
// ===== library: MasterCopy "FB_FIR_LowPass" =====

// folder: UUT/FIR

FUNCTION_BLOCK "FB_FIR_LowPass"   // FB23, SCL
{ S7_Optimized_Access := 'TRUE' }
VERSION : 0.1
   VAR_INPUT
      Enable : Bool;   // filter active
      Reset : Bool;   // restart: the filter is filled with the current X (no start-up ramp)
      X : LReal;   // input sample
      Fc_Set : LReal := 1.0;   // [Hz] requested -3 dB cutoff, about 0.23 Hz ... 20 Hz; a change restarts the filter
      Ts_Limit : LReal := 0.01;   // [s] longer intervals (e.g. a communication peak) are ignored
      Ts_Tol : LReal := 0.05;   // allowed deviation of the average cycle from TS_DESIGN (0.05 = 5 %)
   END_VAR
   VAR_OUTPUT
      Y : LReal;   // filtered output
      M_Act : Int;   // window length of each stage in samples
      Fc_Eff : LReal;   // effective -3 dB cutoff for M_Act and Ts_Meas [Hz]
      Delay : LReal;   // delay of the output (group delay) [s]
      Ts_Meas : LReal;   // average sample period = average OB1 cycle, over about 1 s [s]
      Ts_Valid : Bool;   // TRUE = RUNTIME gave a plausible interval in this call
      Ts_Drift : Bool;   // TRUE = the average cycle differs from TS_DESIGN by more than Ts_Tol: the cutoff is off
   END_VAR
   VAR
      RtMem : LReal;   // memory of RUNTIME
      First : Bool := TRUE;   // first call: no interval yet
      HaveTs : Bool;   // TRUE after the first valid interval
      TsAvg : LReal;   // average of the valid intervals [s]
      Filled : Bool;   // TRUE after the buffers were filled
      "M" : Int;   // window length in use
      Pos : Int;   // ring buffer index: oldest sample of every stage, overwritten in this call
      Sum : Array[0..3] of LReal;   // running sum of every stage
      Buf : Array[0..3, 0..999] of LReal;   // last M inputs of every stage; second bound = M_MAX - 1
   END_VAR
   VAR_TEMP
      tsRaw : LReal;
      mReq : DInt;
      v : LReal;
      s : Int;
      i : Int;
   END_VAR
   VAR CONSTANT
      STAGE_LAST : Int := 3;   // 4 stages
      M_MAX : Int := 1000;   // bound of #Buf: lowest cutoff about 0.23 Hz at 1 ms
      TS_DESIGN : LReal := 0.001;   // design sample period = OB1 cycle [s]
      FC_FACTOR : LReal := 0.2276;   // 4 stages: -3 dB cutoff = FC_FACTOR / (M * Ts)
      TS_SMOOTH : LReal := 0.001;   // weight of a new interval in #TsAvg (about 1000 cycles = 1 s)
   END_VAR
BEGIN

    REGION Description
        // FIR low-pass made of 4 cascaded moving averages of M samples each (4 * (M - 1) + 1 taps, all positive):
        // linear phase, DC gain 1, no overshoot on a step. Every stage keeps a running sum, so one call costs the
        // same for any M: the cutoff can go low without more computing time, only more memory (#Buf).
        //   -3 dB at Fc = 0.2276 / (M * Ts); zeros at multiples of 1 / (M * Ts); everything above the first zero
        //   is damped by at least 53 dB. Delay = 2 * (M - 1) * Ts, about 0.45 / Fc.
        // M follows from Fc_Set and TS_DESIGN (rounded, 1 ... M_MAX), so Fc_Eff differs slightly from Fc_Set.
        // Call in every OB1 cycle and unconditionally: RUNTIME measures the time between two calls.
    END_REGION

    REGION Sample period (RUNTIME: time since the previous call, in seconds)
        #tsRaw := RUNTIME(#RtMem);
        #Ts_Valid := NOT #First AND #tsRaw > 0.0 AND #tsRaw <= #Ts_Limit;
        #First := FALSE;
        IF #Ts_Valid THEN
            IF #HaveTs THEN
                #TsAvg := #TsAvg + (#tsRaw - #TsAvg) * #TS_SMOOTH;
            ELSE
                #TsAvg := #tsRaw;
                #HaveTs := TRUE;
            END_IF;
        END_IF;
        // an invalid interval keeps the last average; before the first valid one: design period
        IF #HaveTs THEN
            #Ts_Meas := #TsAvg;
        ELSE
            #Ts_Meas := #TS_DESIGN;
        END_IF;
        #Ts_Drift := #HaveTs AND ABS(#Ts_Meas - #TS_DESIGN) > #Ts_Tol * #TS_DESIGN;
    END_REGION

    REGION Window length from the requested cutoff
        // LREAL_TO_DINT rounds to the nearest value; below the lowest cutoff: M_MAX (also for Fc_Set <= 0)
        IF #Fc_Set > #FC_FACTOR / (INT_TO_LREAL(#M_MAX) * #TS_DESIGN) THEN
            #mReq := LREAL_TO_DINT(#FC_FACTOR / (#Fc_Set * #TS_DESIGN));
        ELSE
            #mReq := INT_TO_DINT(#M_MAX);
        END_IF;
        IF #mReq < 1 THEN
            #mReq := 1;
        END_IF;
    END_REGION

    REGION Filter
        IF #Reset OR NOT #Filled OR #mReq <> INT_TO_DINT(#M) THEN
            // (re)start: fill every stage with the current input, so the output starts at X
            #M := DINT_TO_INT(#mReq);
            FOR #s := 0 TO #STAGE_LAST DO
                FOR #i := 0 TO #M - 1 DO
                    #Buf[#s, #i] := #X;
                END_FOR;
                #Sum[#s] := #X * INT_TO_LREAL(#M);
            END_FOR;
            #Pos := 0;
            #Filled := TRUE;
            #Y := #X;
        ELSIF #Enable THEN
            #v := #X;
            FOR #s := 0 TO #STAGE_LAST DO
                #Sum[#s] := #Sum[#s] + #v - #Buf[#s, #Pos];   // add the newest, drop the oldest
                #Buf[#s, #Pos] := #v;
                #v := #Sum[#s] / INT_TO_LREAL(#M);   // average of this stage = input of the next one
            END_FOR;
            #Pos := #Pos + 1;
            IF #Pos >= #M THEN
                #Pos := 0;
            END_IF;
            #Y := #v;
        END_IF;

        #M_Act := #M;
        #Fc_Eff := #FC_FACTOR / (INT_TO_LREAL(#M) * #Ts_Meas);
        #Delay := 2.0 * INT_TO_LREAL(#M - 1) * #Ts_Meas;
    END_REGION
END_FUNCTION_BLOCK

// ===== library: MasterCopy "FB_FIR_LP100" =====

// folder: UUT/FIR

FUNCTION_BLOCK "FB_FIR_LP100"   // FB21, SCL
{ S7_Optimized_Access := 'TRUE' }
VERSION : 0.4
   VAR_INPUT
      Enable : Bool;   // filter active
      Reset : Bool;   // clear the delay line
      X : LReal;   // input sample
      Ts_Limit : LReal := 0.01;   // [s] longer intervals (e.g. a communication peak) are ignored
      Ts_Tol : LReal := 0.05;   // allowed deviation of the average cycle from TS_DESIGN (0.05 = 5 %)
   END_VAR
   VAR_OUTPUT
      Y : LReal;   // filtered output
      Ts_Meas : LReal;   // average sample period = average OB1 cycle, over about 1 s [s]
      Ts_Valid : Bool;   // TRUE = RUNTIME gave a plausible interval in this call
      Ts_Drift : Bool;   // TRUE = the average cycle differs from TS_DESIGN by more than Ts_Tol: the cutoff is off
      Fc_Eff : LReal;   // effective -3 dB cutoff for Ts_Meas [Hz]
   END_VAR
   VAR
      RtMem : LReal;   // memory of RUNTIME
      First : Bool := TRUE;   // first call: no interval yet
      HaveTs : Bool;   // TRUE after the first valid interval
      TsAvg : LReal;   // average of the valid intervals [s]
      Pos : Int;   // index of the newest sample in #Line (ring buffer)
      Line : Array[0..16] of LReal;   // delay line (ring buffer)
      Coef : Array[0..16] of LReal;   // [0] [1] [2] [3] [4] [5] [6] [7] [8] [9] [10] [11] [12] [13] [14] [15] [16] filter taps, do not change online
   END_VAR
   VAR_TEMP
      tsRaw : LReal;
      acc : LReal;
      i : Int;
      j : Int;
   END_VAR
   VAR CONSTANT
      LAST_TAP : Int := 16;   // number of taps - 1 = upper bound of #Line and #Coef
      TS_DESIGN : LReal := 0.001;   // design sample period = OB1 cycle [s], fs = 1000 Hz
      FC_DESIGN : LReal := 100.0;   // design -3 dB cutoff [Hz]
      TS_SMOOTH : LReal := 0.001;   // weight of a new interval in #TsAvg (about 1000 cycles = 1 s)
   END_VAR
   // Coef[0] := -1.48651536431772E-19;
   // Coef[1] := -0.000353560113498742;
   // Coef[2] := -0.00350832878720326;
   // Coef[3] := -0.00907130526178393;
   // Coef[4] := -0.00367490473275513;
   // Coef[5] := 0.037817961535658;
   // Coef[6] := 0.124770149738866;
   // Coef[7] := 0.221633438427618;
   // Coef[8] := 0.264773098386197;
   // Coef[9] := 0.221633438427618;
   // Coef[10] := 0.124770149738866;
   // Coef[11] := 0.037817961535658;
   // Coef[12] := -0.00367490473275513;
   // Coef[13] := -0.00907130526178392;
   // Coef[14] := -0.00350832878720326;
   // Coef[15] := -0.000353560113498744;
   // Coef[16] := -1.48651536431772E-19;
BEGIN

    REGION Description
        // FIR low-pass, 17 taps (Blackman-windowed sinc), linear phase, group delay 8 samples = 8 ms, DC gain 1.
        // Designed for an OB1 cycle of 1 ms: -3 dB at 100 Hz, -60 dB from 287 Hz, below -72 dB from 300 Hz to 500 Hz.
        // The taps are fixed, so the cutoff scales with the average cycle: Fc_Eff = 100 Hz * TS_DESIGN / Ts_Meas.
        // Ts_Drift reports a lasting deviation; short peaks of the cycle are averaged out.
        // Call in every OB1 cycle and unconditionally: RUNTIME measures the time between two calls.
    END_REGION

    REGION Sample period (RUNTIME: time since the previous call, in seconds)
        #tsRaw := RUNTIME(#RtMem);
        #Ts_Valid := NOT #First AND #tsRaw > 0.0 AND #tsRaw <= #Ts_Limit;
        #First := FALSE;
        IF #Ts_Valid THEN
            IF #HaveTs THEN
                #TsAvg := #TsAvg + (#tsRaw - #TsAvg) * #TS_SMOOTH;
            ELSE
                #TsAvg := #tsRaw;
                #HaveTs := TRUE;
            END_IF;
        END_IF;
        // an invalid interval keeps the last average; before the first valid one: design period
        IF #HaveTs THEN
            #Ts_Meas := #TsAvg;
        ELSE
            #Ts_Meas := #TS_DESIGN;
        END_IF;
        #Fc_Eff := #FC_DESIGN * #TS_DESIGN / #Ts_Meas;
        #Ts_Drift := #HaveTs AND ABS(#Ts_Meas - #TS_DESIGN) > #Ts_Tol * #TS_DESIGN;
    END_REGION

    REGION Convolution (ring buffer: one write per cycle instead of shifting all samples)
        IF #Reset THEN
            FOR #i := 0 TO #LAST_TAP DO
                #Line[#i] := 0.0;
            END_FOR;
            #Pos := 0;
            #Y := 0.0;
        ELSIF #Enable THEN
            #Pos := #Pos + 1;
            IF #Pos > #LAST_TAP THEN
                #Pos := 0;
            END_IF;
            #Line[#Pos] := #X;
            #acc := 0.0;
            #j := #Pos;   // Coef[i] * sample of i cycles ago
            FOR #i := 0 TO #LAST_TAP DO
                #acc := #acc + #Coef[#i] * #Line[#j];
                #j := #j - 1;
                IF #j < 0 THEN
                    #j := #LAST_TAP;
                END_IF;
            END_FOR;
            #Y := #acc;
        END_IF;
    END_REGION
END_FUNCTION_BLOCK

// ===== library: MasterCopy "UnitTest_FIR_LowPass" =====

// folder: UUT/FIR

FUNCTION_BLOCK "UnitTest_FIR_LowPass"   // FB22, SCL
{ S7_Optimized_Access := 'TRUE' }
VERSION : 0.1
   VAR_INPUT
      reset : Bool;   // TRUE = start the test again (as "DB_UnitTestControl".reset)
   END_VAR
   VAR_OUTPUT
      Done : Bool;   // TRUE when all test steps are finished
   END_VAR
   VAR_IN_OUT
      "Step" : UDInt;   // current step; only increases: 0, 10, 20, 30, 40, 9900
   END_VAR
   VAR
      TestCase : String[24];   // signal of the current step (online monitoring)
      Fir : "FB_FIR_LowPass";   // device under test
      StepTimer : TON_TIME;   // 5 s per signal
      StepRun : Bool;   // FALSE for one cycle after a step change: restarts #StepTimer
      StepSamples : DInt;   // filter calls since the start of the step
      Counting : Bool;   // TRUE = the filter has settled and, for a sine, a signal period has started
      Seed : DWord := 16#2545_F491;   // state of the noise generator (xorshift32), never 0; restarted in step 0
      Sig : Struct   // signal of the current step: X = Offset + Amp * sin(Phase) + noise
         Offset : LReal;
         Amp : LReal;
         K : LReal;   // frequency as a multiple of the effective cutoff: f = K * Fc_Eff
         NoiseAmp : LReal;   // uniform noise in -NoiseAmp ... +NoiseAmp
         FreqHz : LReal;   // resulting frequency (online monitoring)
         Phase : LReal;
         Noise : LReal;
         X : LReal;   // filter input
      END_STRUCT;
      Acc : Struct   // running sums while #Counting
         N : DInt;
         SumY : LReal;
         SumY2 : LReal;
         SumI : LReal;   // Y * sin(Phase)
         SumQ : LReal;   // Y * cos(Phase)
      END_STRUCT;
      Full : Struct   // sums of #Acc at the end of the last whole signal period (sine steps)
         N : DInt;
         SumI : LReal;
         SumQ : LReal;
      END_STRUCT;
      Result : Array[1..4] of Struct   // one entry per signal step: measured value and limits
         Value : LReal;   // step 10: mean of Y; steps 20 ... 40: amplitude of Y at the signal frequency
         Lo : LReal;
         Hi : LReal;
         N : DInt;   // evaluated samples; 0 = the step was too short for an evaluation
         Pass : Bool;
      END_STRUCT;
      NoiseRatio : LReal;   // step 10: standard deviation of Y / standard deviation of the input noise
   END_VAR
   VAR_TEMP
      _ret : Bool;
      res : Int;   // index into #Result
      mean : LReal;
   END_VAR
   VAR CONSTANT
      LAST_STEP : UDInt := 16#FFFF_FFFF;
      STEP_FINISH : UDInt := 9900;
      STEP_TIME : Time := T#5S;   // duration of every signal
      TEST_FC : LReal := 10.0;   // [Hz] cutoff under test: M = 11, so the slow sine of step 20 fits into 5 s
      TWO_PI : LReal := 6.28318530717959;
      NOISE_RATIO_MAX : LReal := 0.3;   // white noise gain of the taps for M = 11 is 0.209
   END_VAR
BEGIN

    REGION BLOCK INFO HEADER
        //===============================================================================
        // Title:            Unit test for FB_FIR_LowPass
        // Comment/Function: Four signals with uniform noise, 5 s each; checks DC gain, noise reduction,
        //                   passband, -3 dB point and stopband at Fc_Set = TEST_FC
        // Requirements:     "FB_FIR_LowPass", unit test framework ("BeforeEach", "AfterEach", "assertTrue",
        //                   "DB_UnitTestControl")
        // Restrictions:     call in every OB1 cycle, unconditionally. The OB1 cycle must be below about 4 ms,
        //                   otherwise 5 s give too few samples (step 10 and step 20 become unreliable)
        //-------------------------------------------------------------------------------
        // Change log table:
        // Version  | Date       | Expert in charge       | Changes applied
        //----------|------------|------------------------|------------------------------
        // 00.00.01 | 21.11.2026 | Roman Butsenko
        //                         First released version, from UnitTest_FIR_LP100 V0.0.3
        //===============================================================================
    END_REGION
    REGION Description
        // Steps (each signal runs STEP_TIME; the evaluation starts after the filter length, 4 * M_Act calls):
        //   10  DC 1.0 + noise 0.5     -> mean of Y 0.98 ... 1.02, noise std reduced below NOISE_RATIO_MAX
        //   20  sine 0.1 * Fc + noise  -> amplitude 0.95 ... 1.05 (passband, theory 0.997)
        //   30  sine 1.0 * Fc + noise  -> amplitude 0.65 ... 0.76 (-3 dB point, theory 0.707)
        //   40  sine 6.6 * Fc + noise  -> amplitude <= 0.004 (stopband, 1.5 x first zero, theory 0.0023 = -53 dB)
        // The filter runs with Fc_Set = TEST_FC; M only scales the filter, so other cutoffs behave the same.
        // Fc is "Fir".Fc_Eff, so the signal has the same frequency per filter call for any OB1 cycle. The amplitude
        // is measured by correlation with sin and cos of the signal phase over whole signal periods, which ignores
        // the noise and the filter delay. Results: #Result[1..4], #NoiseRatio.
    END_REGION

    REGION Reset
        IF "DB_UnitTestControl".reset = 1 OR #reset THEN
            #Done := FALSE;
            #Step := 0;
            #StepRun := FALSE;
            #TestCase := '';
            RETURN;
        END_IF;
    END_REGION

    REGION Signal of this step
        CASE #Step OF
            10:
                #TestCase := 'DC + noise';
                #Sig.Offset := 1.0; #Sig.Amp := 0.0; #Sig.K := 0.0; #Sig.NoiseAmp := 0.5;
            20:
                #TestCase := 'Sine 0.1 Fc + noise';
                #Sig.Offset := 0.0; #Sig.Amp := 1.0; #Sig.K := 0.1; #Sig.NoiseAmp := 0.2;
            30:
                #TestCase := 'Sine 1.0 Fc + noise';
                #Sig.Offset := 0.0; #Sig.Amp := 1.0; #Sig.K := 1.0; #Sig.NoiseAmp := 0.2;
            40:
                #TestCase := 'Sine 6.6 Fc + noise';
                #Sig.Offset := 0.0; #Sig.Amp := 1.0; #Sig.K := 6.6; #Sig.NoiseAmp := 0.2;
            ELSE
                #Sig.Offset := 0.0; #Sig.Amp := 0.0; #Sig.K := 0.0; #Sig.NoiseAmp := 0.0;
        END_CASE;

        // noise: xorshift32, scaled to -NoiseAmp ... +NoiseAmp
        #Seed := #Seed XOR SHL(IN := #Seed, N := 13);
        #Seed := #Seed XOR SHR(IN := #Seed, N := 17);
        #Seed := #Seed XOR SHL(IN := #Seed, N := 5);
        #Sig.Noise := (UDINT_TO_LREAL(DWORD_TO_UDINT(#Seed)) / 4294967296.0 * 2.0 - 1.0) * #Sig.NoiseAmp;
        #Sig.X := #Sig.Offset + #Sig.Amp * SIN(#Sig.Phase) + #Sig.Noise;

        #Fir(Enable := TRUE,
             Reset := #Step = 0,
             X := #Sig.X,
             Fc_Set := #TEST_FC);
        #StepSamples := #StepSamples + 1;

        // step timer: restarts one cycle after every step change
        #StepTimer(IN := #StepRun, PT := #STEP_TIME);
        #StepRun := TRUE;

        // running sums
        IF #Counting THEN
            #Acc.N := #Acc.N + 1;
            #Acc.SumY := #Acc.SumY + #Fir.Y;
            #Acc.SumY2 := #Acc.SumY2 + #Fir.Y * #Fir.Y;
            #Acc.SumI := #Acc.SumI + #Fir.Y * SIN(#Sig.Phase);
            #Acc.SumQ := #Acc.SumQ + #Fir.Y * COS(#Sig.Phase);
        END_IF;

        // next phase: f = K * Fc_Eff; Fc_Eff * Ts_Meas is constant, so the phase step per call is constant
        #Sig.FreqHz := #Sig.K * #Fir.Fc_Eff;
        #Sig.Phase := #Sig.Phase + #TWO_PI * #Sig.FreqHz * #Fir.Ts_Meas;
        IF #Sig.Phase >= #TWO_PI THEN   // a signal period is complete
            #Sig.Phase := #Sig.Phase - #TWO_PI;
            IF #Counting THEN   // keep the sums over whole periods
                #Full.N := #Acc.N;
                #Full.SumI := #Acc.SumI;
                #Full.SumQ := #Acc.SumQ;
            ELSIF #StepSamples >= 4 * INT_TO_DINT(#Fir.M_Act) THEN   // settled: start counting with a new period
                #Counting := TRUE;
            END_IF;
        END_IF;
        IF #Sig.K = 0.0 AND #StepSamples >= 4 * INT_TO_DINT(#Fir.M_Act) THEN   // DC: no periods, count once settled
            #Counting := TRUE;
        END_IF;
    END_REGION

    REGION Test steps
        CASE #Step OF
            0:
                "BeforeEach"(iName := GetBlockName(DINT#16));
                #Result[1].Lo := 0.98;  #Result[1].Hi := 1.02;
                #Result[2].Lo := 0.95;  #Result[2].Hi := 1.05;
                #Result[3].Lo := 0.65;  #Result[3].Hi := 0.76;
                #Result[4].Lo := 0.0;   #Result[4].Hi := 0.004;
                #NoiseRatio := 0.0;
                #Seed := 16#2545_F491;   // same noise in every run, so a failure can be repeated
                #Step := 10;
                #StepRun := FALSE;
                #StepSamples := 0;
                #Counting := FALSE;
                #Sig.Phase := 0.0;
                #Acc.N := 0; #Acc.SumY := 0.0; #Acc.SumY2 := 0.0; #Acc.SumI := 0.0; #Acc.SumQ := 0.0;
                #Full.N := 0; #Full.SumI := 0.0; #Full.SumQ := 0.0;

            10, 20, 30, 40:
                IF #StepTimer.Q THEN
                    #res := UDINT_TO_INT(#Step / 10);
                    #Result[#res].Value := 0.0;
                    IF #Step = 10 THEN
                        #Result[#res].N := #Acc.N;
                        IF #Acc.N > 0 THEN
                            #mean := #Acc.SumY / DINT_TO_LREAL(#Acc.N);
                            #Result[#res].Value := #mean;
                            // std of Y / std of the input noise (uniform: NoiseAmp / sqrt(3))
                            #NoiseRatio := SQRT(MAX(IN1 := #Acc.SumY2 / DINT_TO_LREAL(#Acc.N) - #mean * #mean, IN2 := 0.0))
                                           / (#Sig.NoiseAmp / SQRT(3.0));
                            #_ret := "assertTrue"(#NoiseRatio <= #NOISE_RATIO_MAX);   // noise is reduced
                        END_IF;
                    ELSE
                        #Result[#res].N := #Full.N;
                        IF #Full.N > 0 THEN
                            #Result[#res].Value := 2.0 / DINT_TO_LREAL(#Full.N) * SQRT(#Full.SumI * #Full.SumI + #Full.SumQ * #Full.SumQ);
                        END_IF;
                    END_IF;
                    #Result[#res].Pass := #Result[#res].N > 0 AND #Result[#res].Value >= #Result[#res].Lo AND #Result[#res].Value <= #Result[#res].Hi;
                    #_ret := "assertTrue"(#Result[#res].Pass);

                    // next signal
                    IF #Step < 40 THEN
                        #Step := #Step + 10;
                    ELSE
                        #Step := #STEP_FINISH;
                    END_IF;
                    #StepRun := FALSE;
                    #StepSamples := 0;
                    #Counting := FALSE;
                    #Sig.Phase := 0.0;
                    #Acc.N := 0; #Acc.SumY := 0.0; #Acc.SumY2 := 0.0; #Acc.SumI := 0.0; #Acc.SumQ := 0.0;
                    #Full.N := 0; #Full.SumI := 0.0; #Full.SumQ := 0.0;
                END_IF;

            #STEP_FINISH: // all test steps are done
                #Done := TRUE;
                "AfterEach"();
                #Step := #LAST_STEP;

            #LAST_STEP:
                // just idle
                ;

            ELSE // step number without a label: report it and finish the test
                #_ret := "assertTrue"(FALSE);
                #Step := #STEP_FINISH;
        END_CASE;
    END_REGION
END_FUNCTION_BLOCK

// ===== library: MasterCopy "UnitTest_FIR_LP100" =====

// folder: UUT/FIR

FUNCTION_BLOCK "UnitTest_FIR_LP100"   // FB20, SCL
{ S7_Optimized_Access := 'TRUE' }
VERSION : 0.3
   VAR_INPUT
      reset : Bool;   // TRUE = start the test again (as "DB_UnitTestControl".reset)
   END_VAR
   VAR_OUTPUT
      Done : Bool;   // TRUE when all test steps are finished
   END_VAR
   VAR_IN_OUT
      "Step" : UDInt;   // current step; only increases: 0, 10, 20, 30, 40, 9900
   END_VAR
   VAR
      TestCase : String[24];   // signal of the current step (online monitoring)
      Fir : "FB_FIR_LP100";   // device under test
      StepTimer : TON_TIME;   // 5 s per signal
      StepRun : Bool;   // FALSE for one cycle after a step change: restarts #StepTimer
      StepSamples : DInt;   // filter calls since the start of the step
      Counting : Bool;   // TRUE = the filter has settled and, for a sine, a signal period has started
      Seed : DWord := 16#2545_F491;   // state of the noise generator (xorshift32), never 0; restarted in step 0
      Sig : Struct   // signal of the current step: X = Offset + Amp * sin(Phase) + noise
         Offset : LReal;
         Amp : LReal;
         K : LReal;   // frequency as a multiple of the effective cutoff: f = K * Fc_Eff
         NoiseAmp : LReal;   // uniform noise in -NoiseAmp ... +NoiseAmp
         FreqHz : LReal;   // resulting frequency (online monitoring)
         Phase : LReal;
         Noise : LReal;
         X : LReal;   // filter input
      END_STRUCT;
      Acc : Struct   // running sums while #Counting
         N : DInt;
         SumY : LReal;
         SumY2 : LReal;
         SumI : LReal;   // Y * sin(Phase)
         SumQ : LReal;   // Y * cos(Phase)
      END_STRUCT;
      Full : Struct   // sums of #Acc at the end of the last whole signal period (sine steps)
         N : DInt;
         SumI : LReal;
         SumQ : LReal;
      END_STRUCT;
      Result : Array[1..4] of Struct   // one entry per signal step: measured value and limits
         Value : LReal;   // step 10: mean of Y; steps 20 ... 40: amplitude of Y at the signal frequency
         Lo : LReal;
         Hi : LReal;
         N : DInt;   // evaluated samples; 0 = the step was too short for an evaluation
         Pass : Bool;
      END_STRUCT;
      NoiseRatio : LReal;   // step 10: standard deviation of Y / standard deviation of the input noise
   END_VAR
   VAR_TEMP
      _ret : Bool;
      res : Int;   // index into #Result
      mean : LReal;
   END_VAR
   VAR CONSTANT
      LAST_STEP : UDInt := 16#FFFF_FFFF;
      STEP_FINISH : UDInt := 9900;
      STEP_TIME : Time := T#5S;   // duration of every signal
      SETTLE_SAMPLES : DInt := 17;   // filter calls before the evaluation starts (= number of taps)
      TWO_PI : LReal := 6.28318530717959;
      NOISE_RATIO_MAX : LReal := 0.55;   // white noise gain of the taps is 0.450
   END_VAR
BEGIN

    REGION BLOCK INFO HEADER
        //===============================================================================
        // Title:            Unit test for FB_FIR_LP100
        // Comment/Function: Four signals with uniform noise, 5 s each; checks DC gain, noise reduction,
        //                   passband, -3 dB point and stopband
        // Requirements:     "FB_FIR_LP100", unit test framework ("BeforeEach", "AfterEach", "assertTrue",
        //                   "DB_UnitTestControl")
        // Restrictions:     call in every OB1 cycle, unconditionally. The OB1 cycle must be below about 10 ms,
        //                   otherwise 5 s give too few samples (step 10 and step 20 become unreliable)
        //-------------------------------------------------------------------------------
        // Change log table:
        // Version  | Date       | Expert in charge       | Changes applied
        //----------|------------|------------------------|------------------------------
        // 00.00.01 | 21.11.2026 | Roman Butsenko
        //                         First released version
        // 00.00.02 | 21.11.2026 | Roman Butsenko
        //                         Step as InOut; OB1 instead of a cyclic OB; noise restarts in step 0;
        //                         sine amplitude over whole signal periods; settling counted in filter calls
        // 00.00.03 | 21.11.2026 | Roman Butsenko
        //                         17 taps for a 1 ms OB1 cycle: settling 17 calls, noise limit 0.55,
        //                         stopband test at 3 Fc (5 Fc = 500 Hz is the Nyquist frequency at 1 ms)
        //===============================================================================
    END_REGION
    REGION Description
        // Steps (each signal runs STEP_TIME; the evaluation starts SETTLE_SAMPLES calls after the step change):
        //   10  DC 1.0 + noise 0.5     -> mean of Y 0.98 ... 1.02, noise std reduced below NOISE_RATIO_MAX
        //   20  sine 0.1 * Fc + noise  -> amplitude 0.95 ... 1.05 (passband, theory 0.997)
        //   30  sine 1.0 * Fc + noise  -> amplitude 0.65 ... 0.76 (-3 dB point, theory 0.707)
        //   40  sine 3.0 * Fc + noise  -> amplitude <= 0.001 (stopband, theory 0.00024 = -73 dB)
        // Fc is "Fir".Fc_Eff, so the signal has the same frequency per filter call for any OB1 cycle. The amplitude
        // is measured by correlation with sin and cos of the signal phase over whole signal periods, which ignores
        // the noise and the filter delay. Results: #Result[1..4], #NoiseRatio.
    END_REGION

    REGION Reset
        IF "DB_UnitTestControl".reset = 1 OR #reset THEN
            #Done := FALSE;
            #Step := 0;
            #StepRun := FALSE;
            #TestCase := '';
            RETURN;
        END_IF;
    END_REGION

    REGION Signal of this step
        CASE #Step OF
            10:
                #TestCase := 'DC + noise';
                #Sig.Offset := 1.0; #Sig.Amp := 0.0; #Sig.K := 0.0; #Sig.NoiseAmp := 0.5;
            20:
                #TestCase := 'Sine 0.1 Fc + noise';
                #Sig.Offset := 0.0; #Sig.Amp := 1.0; #Sig.K := 0.1; #Sig.NoiseAmp := 0.2;
            30:
                #TestCase := 'Sine 1.0 Fc + noise';
                #Sig.Offset := 0.0; #Sig.Amp := 1.0; #Sig.K := 1.0; #Sig.NoiseAmp := 0.2;
            40:
                #TestCase := 'Sine 3.0 Fc + noise';
                #Sig.Offset := 0.0; #Sig.Amp := 1.0; #Sig.K := 3.0; #Sig.NoiseAmp := 0.2;
            ELSE
                #Sig.Offset := 0.0; #Sig.Amp := 0.0; #Sig.K := 0.0; #Sig.NoiseAmp := 0.0;
        END_CASE;

        // noise: xorshift32, scaled to -NoiseAmp ... +NoiseAmp
        #Seed := #Seed XOR SHL(IN := #Seed, N := 13);
        #Seed := #Seed XOR SHR(IN := #Seed, N := 17);
        #Seed := #Seed XOR SHL(IN := #Seed, N := 5);
        #Sig.Noise := (UDINT_TO_LREAL(DWORD_TO_UDINT(#Seed)) / 4294967296.0 * 2.0 - 1.0) * #Sig.NoiseAmp;
        #Sig.X := #Sig.Offset + #Sig.Amp * SIN(#Sig.Phase) + #Sig.Noise;

        #Fir(Enable := TRUE,
             Reset := #Step = 0,
             X := #Sig.X);
        #StepSamples := #StepSamples + 1;

        // step timer: restarts one cycle after every step change
        #StepTimer(IN := #StepRun, PT := #STEP_TIME);
        #StepRun := TRUE;

        // running sums
        IF #Counting THEN
            #Acc.N := #Acc.N + 1;
            #Acc.SumY := #Acc.SumY + #Fir.Y;
            #Acc.SumY2 := #Acc.SumY2 + #Fir.Y * #Fir.Y;
            #Acc.SumI := #Acc.SumI + #Fir.Y * SIN(#Sig.Phase);
            #Acc.SumQ := #Acc.SumQ + #Fir.Y * COS(#Sig.Phase);
        END_IF;

        // next phase: f = K * Fc_Eff; Fc_Eff * Ts_Meas is constant, so the phase step per call is constant
        #Sig.FreqHz := #Sig.K * #Fir.Fc_Eff;
        #Sig.Phase := #Sig.Phase + #TWO_PI * #Sig.FreqHz * #Fir.Ts_Meas;
        IF #Sig.Phase >= #TWO_PI THEN   // a signal period is complete
            #Sig.Phase := #Sig.Phase - #TWO_PI;
            IF #Counting THEN   // keep the sums over whole periods
                #Full.N := #Acc.N;
                #Full.SumI := #Acc.SumI;
                #Full.SumQ := #Acc.SumQ;
            ELSIF #StepSamples >= #SETTLE_SAMPLES THEN   // settled: start counting with a new period
                #Counting := TRUE;
            END_IF;
        END_IF;
        IF #Sig.K = 0.0 AND #StepSamples >= #SETTLE_SAMPLES THEN   // DC: no periods, count once settled
            #Counting := TRUE;
        END_IF;
    END_REGION

    REGION Test steps
        CASE #Step OF
            0:
                "BeforeEach"(iName := GetBlockName(DINT#16));
                #Result[1].Lo := 0.98;  #Result[1].Hi := 1.02;
                #Result[2].Lo := 0.95;  #Result[2].Hi := 1.05;
                #Result[3].Lo := 0.65;  #Result[3].Hi := 0.76;
                #Result[4].Lo := 0.0;   #Result[4].Hi := 0.001;
                #NoiseRatio := 0.0;
                #Seed := 16#2545_F491;   // same noise in every run, so a failure can be repeated
                #Step := 10;
                #StepRun := FALSE;
                #StepSamples := 0;
                #Counting := FALSE;
                #Sig.Phase := 0.0;
                #Acc.N := 0; #Acc.SumY := 0.0; #Acc.SumY2 := 0.0; #Acc.SumI := 0.0; #Acc.SumQ := 0.0;
                #Full.N := 0; #Full.SumI := 0.0; #Full.SumQ := 0.0;

            10, 20, 30, 40:
                IF #StepTimer.Q THEN
                    #res := UDINT_TO_INT(#Step / 10);
                    #Result[#res].Value := 0.0;
                    IF #Step = 10 THEN
                        #Result[#res].N := #Acc.N;
                        IF #Acc.N > 0 THEN
                            #mean := #Acc.SumY / DINT_TO_LREAL(#Acc.N);
                            #Result[#res].Value := #mean;
                            // std of Y / std of the input noise (uniform: NoiseAmp / sqrt(3))
                            #NoiseRatio := SQRT(MAX(IN1 := #Acc.SumY2 / DINT_TO_LREAL(#Acc.N) - #mean * #mean, IN2 := 0.0))
                                           / (#Sig.NoiseAmp / SQRT(3.0));
                            #_ret := "assertTrue"(#NoiseRatio <= #NOISE_RATIO_MAX);   // noise is reduced
                        END_IF;
                    ELSE
                        #Result[#res].N := #Full.N;
                        IF #Full.N > 0 THEN
                            #Result[#res].Value := 2.0 / DINT_TO_LREAL(#Full.N) * SQRT(#Full.SumI * #Full.SumI + #Full.SumQ * #Full.SumQ);
                        END_IF;
                    END_IF;
                    #Result[#res].Pass := #Result[#res].N > 0 AND #Result[#res].Value >= #Result[#res].Lo AND #Result[#res].Value <= #Result[#res].Hi;
                    #_ret := "assertTrue"(#Result[#res].Pass);

                    // next signal
                    IF #Step < 40 THEN
                        #Step := #Step + 10;
                    ELSE
                        #Step := #STEP_FINISH;
                    END_IF;
                    #StepRun := FALSE;
                    #StepSamples := 0;
                    #Counting := FALSE;
                    #Sig.Phase := 0.0;
                    #Acc.N := 0; #Acc.SumY := 0.0; #Acc.SumY2 := 0.0; #Acc.SumI := 0.0; #Acc.SumQ := 0.0;
                    #Full.N := 0; #Full.SumI := 0.0; #Full.SumQ := 0.0;
                END_IF;

            #STEP_FINISH: // all test steps are done
                #Done := TRUE;
                "AfterEach"();
                #Step := #LAST_STEP;

            #LAST_STEP:
                // just idle
                ;

            ELSE // step number without a label: report it and finish the test
                #_ret := "assertTrue"(FALSE);
                #Step := #STEP_FINISH;
        END_CASE;
    END_REGION
END_FUNCTION_BLOCK